// Public HMI interface for fb_CamCoupler - the struct an HMI binds.
// No HMIbaseDevice: fb_CamCoupler is standalone and does NOT extend abs_fb_Device.
TYPE ST_CamCoupler_HMI_Interface :
STRUCT
    Status   : ST_CamCoupler_HMI_Status;
    Commands : ST_CamCoupler_HMI_Commands;
    Config   : ST_CamCoupler_HMI_Config;
END_STRUCT
END_TYPE

(* stored: Version 1.1.0.1
   DUT ST_CamCoupler_HMI_Interface: Id {d1543ff0-d085-4af3-bb9e-aa7c8114f94a} *)
